Staubli VAL3: _tCycleCtrl.pgx

program _tCycleCtrl()
  local bool l_bAckAlarm
  local bool l_bEndCmd
  local bool l_bErr
  local bool l_bHoldCmd
  local bool l_bPowerOff
  local bool l_bPowerOn
  local bool l_bResetCmd
  local bool l_bResetIO
  local bool l_bStartCmd
  local bool l_bStopCmd
  local num l_n
  local bool l_bResult
begin
  //启动程序
  if rs:bToStartCycle and rs:bIsReady
    rs:bToStartCycle=false
    taskCreate "cycle",100,_productCycle()
    wait(taskStatus("cycle")>-1)
  endIf
  //停止程序
  if(rs:bToStopCycle or rs:bIsEstop) and rs:bIsCycle
    rs:bToStopCycle=false
    resetMotion()
    stopMove()
    taskKill("cycle")
    wait(taskStatus("cycle")==-1)
  endIf
  //暂停程序
  if((rs:bToPause) and rs:bIsCycle) or taskStatus("cycle")>1
    rs:bToPause=false
    stopMove()
    rs:bIsPause=true
  endIf
  //暂停恢复程序
  if rs:bIsPause and rs:bIsCycle and rs:bToStartCycle
    rs:bToStartCycle=false
    rs:bIsPause=false
    if !isPowered()
      enablePower()
      l_bResult=watch(isPowered(),1)
      if !l_bResult
        logMsg("恢复生产任务上电超时")
        return
      endIf

    endIf
    autoConnectMove(true)
    restartMove()
  endIf
end
